(* IEC 61131-3 sources: llm-plc-st-eval/data/processed_definitivo/qwen2.5-coder_14b/I6/zero_shot, 3 files *)

(* ---- ejec_1.st ---- *)
FUNCTION_BLOCK FB_Temperatura
VAR_INPUT
    rawTemp : INT;  // Entrada de temperatura cruda (0-27648)
END_VAR

VAR_OUTPUT
    tempC : REAL;   // Temperatura en grados Celsius (0.0-100.0)
    enfriador : BOOL;  // Estado del enfriador (TRUE/FALSE)
    almSensor : BOOL;  // Alarma del sensor (TRUE/FALSE)
END_VAR

VAR
    tempCPrev : REAL;  // Valor previo de temperatura en Celsius
    enfriadorPrev : BOOL;  // Estado previo del enfriador
END_VAR

// Calculo de la temperatura en Celsius
IF rawTemp >= 0 AND rawTemp <= 27648 THEN
    tempC := rawTemp * 100.0 / 27648.0;
    almSensor := FALSE;
ELSE
    tempC := 0.0;
    almSensor := TRUE;
END_IF;

// Control del enfriador con histéresis
IF tempC >= 80.0 THEN
    enfriador := TRUE;
ELSIF tempC <= 75.0 THEN
    enfriador := FALSE;
ELSE
    enfriador := enfriadorPrev;  // Mantener el estado anterior si está en el rango de histéresis
END_IF;

// Actualizar el estado previo del enfriador
enfriadorPrev := enfriador;

END_FUNCTION_BLOCK

(* ---- ejec_2.st ---- *)
FUNCTION_BLOCK FB_Temperatura
VAR_INPUT
    rawTemp : INT; // Entrada de temperatura cruda (0 a 27648)
END_VAR

VAR_OUTPUT
    tempC : REAL; // Temperatura en grados Celsius (0.0 a 100.0)
    enfriador : BOOL; // Estado del enfriador (TRUE: activado, FALSE: desactivado)
    almSensor : BOOL; // Estado de la alarma del sensor (TRUE: activada, FALSE: desactivada)
END_VAR

VAR
    tempCPrev : REAL; // Temperatura anterior para la histéresis
    enfriadorPrev : BOOL; // Estado anterior del enfriador para la histéresis
END_VAR

// Calculo de la temperatura en grados Celsius
IF rawTemp < 0 OR rawTemp > 27648 THEN
    tempC := 0.0;
    almSensor := TRUE;
    enfriador := FALSE;
ELSE
    tempC := rawTemp / 276.48;
    almSensor := FALSE;

    // Control del enfriador con histéresis
    IF tempC >= 80.0 THEN
        enfriador := TRUE;
    ELSIF tempC <= 75.0 THEN
        enfriador := FALSE;
    ELSE
        enfriador := enfriadorPrev; // Mantener el estado anterior
    END_IF
END_IF

// Actualizar el estado anterior del enfriador
enfriadorPrev := enfriador;

(* ---- ejec_3.st ---- *)
FUNCTION_BLOCK FB_Temperatura
VAR_INPUT
    rawTemp : INT; // Entrada de temperatura cruda (0 a 27648)
END_VAR

VAR_OUTPUT
    tempC : REAL; // Temperatura en grados Celsius (0.0 a 100.0)
    enfriador : BOOL; // Estado del enfriador (TRUE: activado, FALSE: desactivado)
    almSensor : BOOL; // Estado de la alarma del sensor (TRUE: activada, FALSE: desactivada)
END_VAR

VAR
    tempCPrev : REAL; // Temperatura anterior para la histéresis
    enfriadorPrev : BOOL; // Estado anterior del enfriador para la histéresis
END_VAR

// Calcula la temperatura en grados Celsius
IF rawTemp < 0 OR rawTemp > 27648 THEN
    tempC := 0.0;
    almSensor := TRUE;
    enfriador := FALSE;
ELSE
    tempC := rawTemp / 276.48; // Conversión de 0-27648 a 0.0-100.0 grados Celsius
    almSensor := FALSE;

    // Control del enfriador con histéresis
    IF tempC >= 80.0 THEN
        enfriador := TRUE;
    ELSIF tempC <= 75.0 THEN
        enfriador := FALSE;
    ELSE
        enfriador := enfriadorPrev; // Mantener el estado anterior si está en la zona de histéresis
    END_IF
END_IF

// Actualiza el estado anterior del enfriador
enfriadorPrev := enfriador;
